TYPE "ST_ProductionUnitParCfg"
VERSION : 0.1
   STRUCT
      SchemaVersion : UInt := 4;
      Timeout : Time := T#8S;
      Preset : DInt := 10;
      IdealCycleMs : UDInt := 1000;
      BaselineMs : UDInt := 1000;
   END_STRUCT;

END_TYPE

